(* PLC project zarechnaya.project, CODESYS CODESYS V3.5 SP17 Patch 3 *)
(* stored: creationDateTime 2026-10-20T05:42:22.3807229, modificationDateTime 1601-01-01T03:00:00 *)

TYPE E_FilterMode : (Off := 0, Filter := 1, Backwash := 2);
END_TYPE
